(* Logix 5000 project; controller TFF vendor 1 type 14 code 107 rev 33.11; software revision 33.04; part 16 of 38 *)
(* tags used below, declared in another part *)
   AddressTotalizer : DINT;   // Temp Address used in modPhaseTotal
   Index : DINT;   // Index
   PLCDST : SINT;   // Current PLC Day Light Saving
   PLCTimeZoneString : STRING;   // Current PLC TimeZone
   TimeZoneUTC0 : STRING;   // String value for Time zone UTC 0
   AnalogPoint : AnalogInput[50];   // Analog Input Array
   Concentration : Concentration;
   ControlLoop_PCV101 : ALIAS FOR ControlLoop[3];
   ControlLoop_PCV101_5ms : ALIAS FOR ControlLoop[4];
   ControlLoop_PCV101_RAMP_OUT : REAL;   // Ramp Output
   Diafiltration : Diafiltration;
   FI201 : ALIAS FOR AnalogPoint[2];
   FQ_Conc : ALIAS FOR Totalizer[0];   // Concentration Totalizer
   FQ_Diaf : ALIAS FOR Totalizer[1];   // DiafiltrationTotalizer
   MiscREAL : REAL[50];   // Misc Real Values
   PCDateTime : DINT[7];   // Date/Time Array from PC
   PCV101 : ALIAS FOR AnalogPoint[3];
   PCV101_Control : PCV_Control;   // PCV101 Control UDT
   PCV101_PID : PCV;   // PCV101 PID Management
   Phase : Phases[6];   // Phase Control Array
   PhaseTotalizer : PhaseTotalizer[18];   // Phase Totalizers Array
   Rack_Murr_Node1_TFF20 : IO_Station;   // Status of Node 1 TFF20
   Rack_Murr_Node1_TFF40 : IO_Station;   // Status of Node 1 TFF40
   Rack_Murr_Node1_TFF80 : IO_Station;   // Status of Node 1 TFF80
   RawAnalogInputArray : INT[50];   // Array of analog input raw
   SysControl : SysControl;   // General system status and command
   ThisSystem : SystemType;
   TimerControl : TimerControl;   // Timer Control
   Timers : Timers[22];   // Timer Array
   Totalizer : Totalizers[20];   // Totalizers Array
   Valve : Valve[100];   // Valve Array
(* MainProgram, continued *)

ROUTINE modPhaseTotal   (* ladder *)
// Phase Totalizer Module
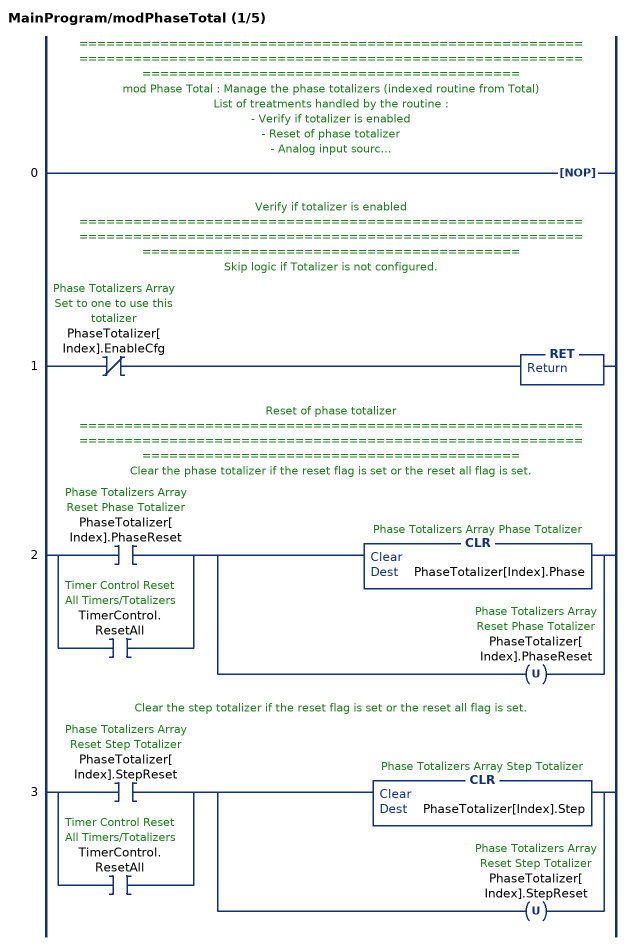
   // ==========================================================================================================================================================
   //                                                                                                   mod Phase Total : Manage the phase totalizers (indexed routine from Total)
   //                                                     List of treatments handled by the routine :
   //                                                          - Verify if totalizer is enabled
   //                                                          - Reset of phase totalizer
   //                                                          - Analog input source
   //                                                          - Calculating the totalizer values
   //                                                     -----------------------------------------------------------------------------------------------------------------------------------------------------
   //                                                     History
   // 		2019-DEC-24 - Merck - Q. Spindler - Initial version for Candidate Release 1.00.00.00.a
   // ==========================================================================================================================================================
   0: NOP();
   // Verify if totalizer is enabled
   // ==========================================================================================================================================================
   // Skip logic if Totalizer is not configured.
   1: XIO(PhaseTotalizer[Index].EnableCfg)RET();
   // Reset of phase totalizer
   // ==========================================================================================================================================================
   // Clear the phase totalizer if the reset flag is set or the reset all flag is set.
   2: [XIC(PhaseTotalizer[Index].PhaseReset) ,XIC(TimerControl.ResetAll) ][CLR(PhaseTotalizer[Index].Phase) ,OTU(PhaseTotalizer[Index].PhaseReset) ];
   // Clear the step totalizer if the reset flag is set or the reset all flag is set.
   3: [XIC(PhaseTotalizer[Index].StepReset) ,XIC(TimerControl.ResetAll) ][CLR(PhaseTotalizer[Index].Step) ,OTU(PhaseTotalizer[Index].StepReset) ];
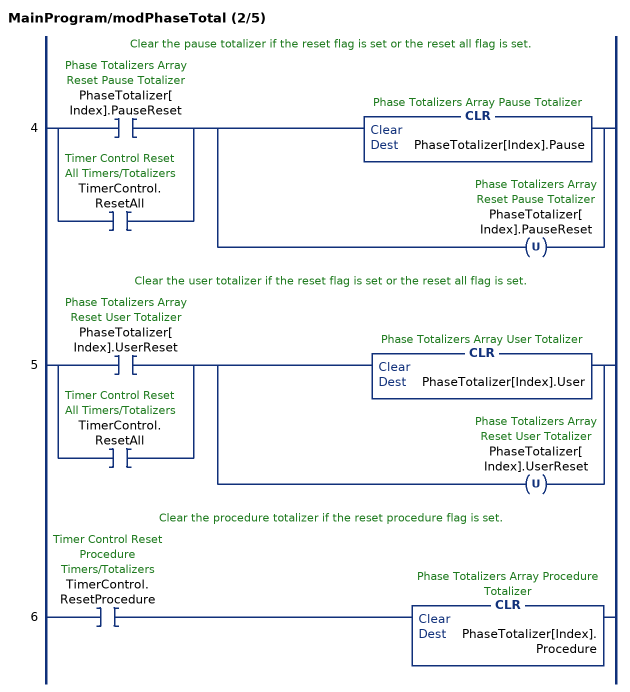
   // Clear the pause totalizer if the reset flag is set or the reset all flag is set.
   4: [XIC(PhaseTotalizer[Index].PauseReset) ,XIC(TimerControl.ResetAll) ][CLR(PhaseTotalizer[Index].Pause) ,OTU(PhaseTotalizer[Index].PauseReset) ];
   // Clear the user totalizer if the reset flag is set or the reset all flag is set.
   5: [XIC(PhaseTotalizer[Index].UserReset) ,XIC(TimerControl.ResetAll) ][CLR(PhaseTotalizer[Index].User) ,OTU(PhaseTotalizer[Index].UserReset) ];
   // Clear the procedure totalizer if the reset procedure flag is set.
   6: XIC(TimerControl.ResetProcedure)CLR(PhaseTotalizer[Index].Procedure);
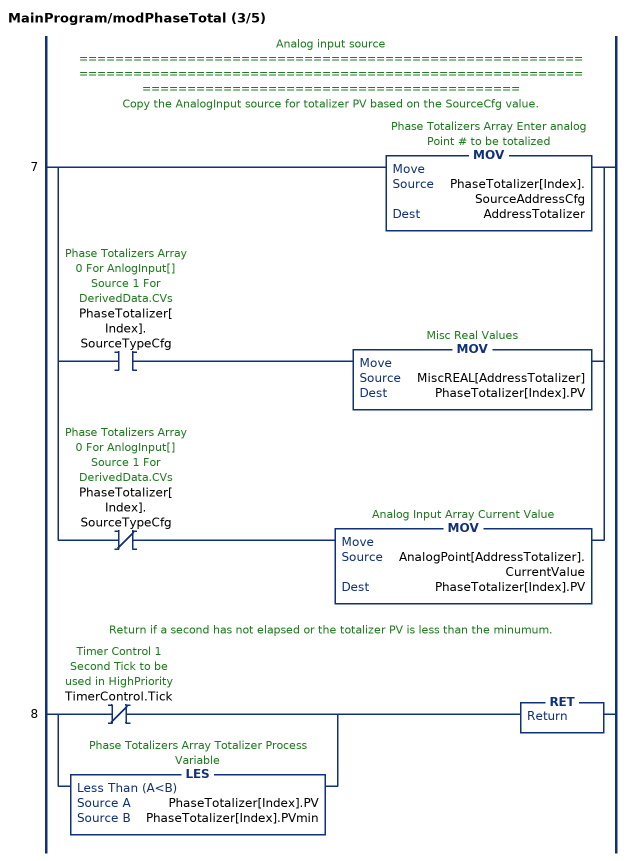
   // Analog input source
   // ==========================================================================================================================================================
   // Copy the AnalogInput source for totalizer PV based on the SourceCfg value.
   7: [MOV(PhaseTotalizer[Index].SourceAddressCfg,AddressTotalizer) ,XIC(PhaseTotalizer[Index].SourceTypeCfg) MOV(MiscREAL[AddressTotalizer],PhaseTotalizer[Index].PV) ,XIO(PhaseTotalizer[Index].SourceTypeCfg) MOV(AnalogPoint[AddressTotalizer].CurrentValue,PhaseTotalizer[Index].PV) ];
   // Return if a second has not elapsed or the totalizer PV is less than the minumum.
   8: [XIO(TimerControl.Tick) ,LES(PhaseTotalizer[Index].PV,PhaseTotalizer[Index].PVmin) ]RET();
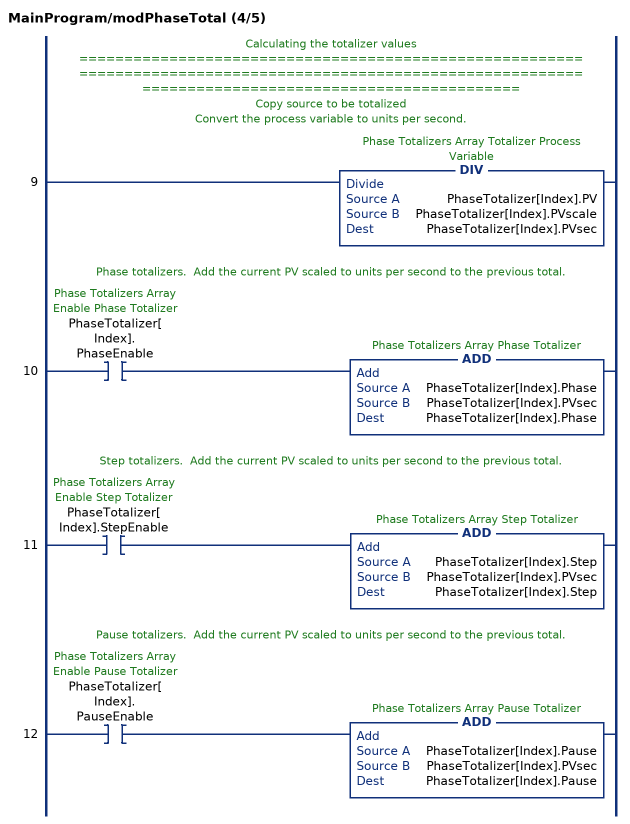
   // Calculating the totalizer values
   // ==========================================================================================================================================================
   // Copy source to be totalized
   // Convert the process variable to units per second.
   9: DIV(PhaseTotalizer[Index].PV,PhaseTotalizer[Index].PVscale,PhaseTotalizer[Index].PVsec);
   // Phase totalizers.  Add the current PV scaled to units per second to the previous total.
   10: XIC(PhaseTotalizer[Index].PhaseEnable)ADD(PhaseTotalizer[Index].Phase,PhaseTotalizer[Index].PVsec,PhaseTotalizer[Index].Phase);
   // Step totalizers.  Add the current PV scaled to units per second to the previous total.
   11: XIC(PhaseTotalizer[Index].StepEnable)ADD(PhaseTotalizer[Index].Step,PhaseTotalizer[Index].PVsec,PhaseTotalizer[Index].Step);
   // Pause totalizers.  Add the current PV scaled to units per second to the previous total.
   12: XIC(PhaseTotalizer[Index].PauseEnable)ADD(PhaseTotalizer[Index].Pause,PhaseTotalizer[Index].PVsec,PhaseTotalizer[Index].Pause);
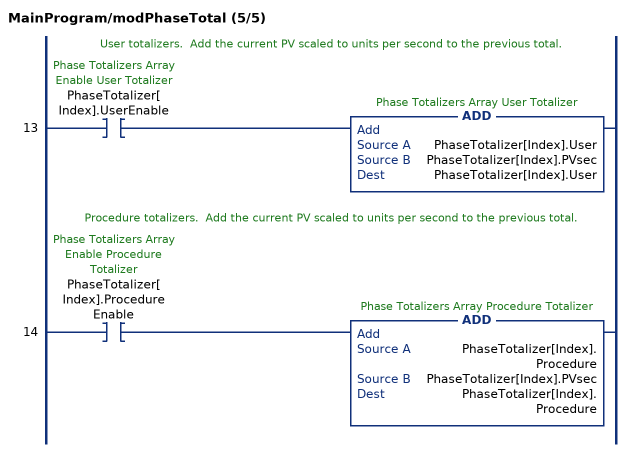
   // User totalizers.  Add the current PV scaled to units per second to the previous total.
   13: XIC(PhaseTotalizer[Index].UserEnable)ADD(PhaseTotalizer[Index].User,PhaseTotalizer[Index].PVsec,PhaseTotalizer[Index].User);
   // Procedure totalizers.  Add the current PV scaled to units per second to the previous total.
   14: XIC(PhaseTotalizer[Index].ProcedureEnable)ADD(PhaseTotalizer[Index].Procedure,PhaseTotalizer[Index].PVsec,PhaseTotalizer[Index].Procedure);
END_ROUTINE

ROUTINE modTotal   (* ladder *)
// Totalizer Module
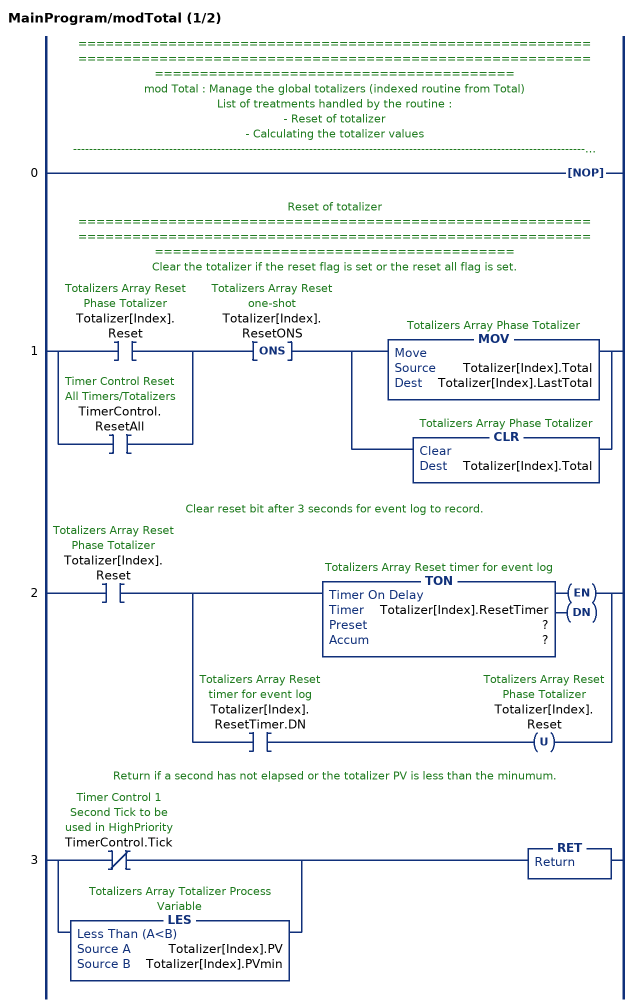
   // ==========================================================================================================================================================
   //                                                                                                   mod Total : Manage the global totalizers (indexed routine from Total)
   //                                                     List of treatments handled by the routine :
   //                                                          - Reset of totalizer
   //                                                          - Calculating the totalizer values
   //                                                     -----------------------------------------------------------------------------------------------------------------------------------------------------
   //                                                     History
   // 		2019-DEC-24 - Merck - Q. Spindler - Initial version for Candidate Release 1.00.00.00.a
   // ==========================================================================================================================================================
   0: NOP();
   // Reset of totalizer
   // ==========================================================================================================================================================
   // Clear the totalizer if the reset flag is set or the reset all flag is set.
   1: [XIC(Totalizer[Index].Reset) ,XIC(TimerControl.ResetAll) ]ONS(Totalizer[Index].ResetONS)[MOV(Totalizer[Index].Total,Totalizer[Index].LastTotal) ,CLR(Totalizer[Index].Total) ];
   // Clear reset bit after 3 seconds for event log to record.
   2: XIC(Totalizer[Index].Reset)[TON(Totalizer[Index].ResetTimer,?,?) ,XIC(Totalizer[Index].ResetTimer.DN) OTU(Totalizer[Index].Reset) ];
   // Return if a second has not elapsed or the totalizer PV is less than the minumum.
   3: [XIO(TimerControl.Tick) ,LES(Totalizer[Index].PV,Totalizer[Index].PVmin) ]RET();
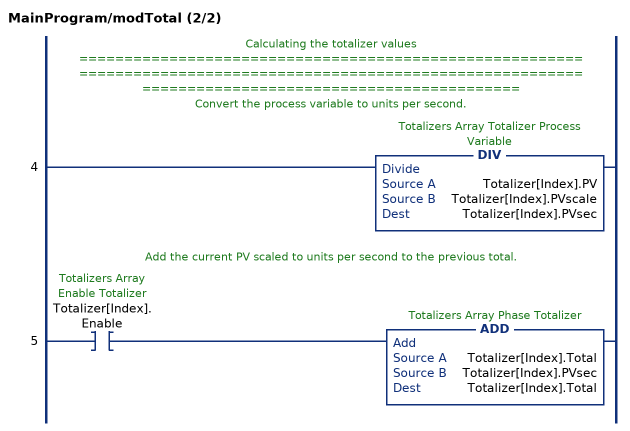
   // Calculating the totalizer values
   // ==========================================================================================================================================================
   // Convert the process variable to units per second.
   4: DIV(Totalizer[Index].PV,Totalizer[Index].PVscale,Totalizer[Index].PVsec);
   // Add the current PV scaled to units per second to the previous total.
   5: XIC(Totalizer[Index].Enable)ADD(Totalizer[Index].Total,Totalizer[Index].PVsec,Totalizer[Index].Total);
END_ROUTINE

ROUTINE PCDateTime   (* structured text *)
   (* =======================================================================
   	PCDateTime : Synchronize the PLC with PC clock
   
   	List of treatments
   		- Synchronization
   
   -----------------------------------------------------------------------------------------------------------------------------------------------------
   	History
   		2019-DEC-24 - Merck - Q. Spindler - Initial version for Candidate Release 1.00.00.00.a
   =========================================================================*)
   
   
   (* Synchronization
   =========================================================================*)
   (*Update the internal PLC clock with the PC clock when the microseconds value is not -1*)
   IF PCDateTime[6] <> -1 THEN;
   	SSV (WALLCLOCKTIME, , DateTime, PCDateTime[0]);
   	PCDateTime[6] := -1;
   END_IF;
   
   (*Get PLC DST settings and set it to 0 of not already*)
   GSV (WALLCLOCKTIME, ,ApplyDST , PLCDST);
   IF PLCDST <> 0 THEN;
   	PLCDST := 0;
   	SSV (WALLCLOCKTIME, ,ApplyDST , PLCDST);
   END_IF;
   
   (*Get PLC TimeZone and set it to UTC0 of not already*)
   GSV (WALLCLOCKTIME, ,TimeZoneString, PLCTimeZoneString);
   IF PLCTimeZoneString <> TimeZoneUTC0 THEN;
   	SSV (WALLCLOCKTIME, ,TimeZoneString , TimeZoneUTC0);
   END_IF;
   
END_ROUTINE

ROUTINE Time   (* ladder *)
// Timekeeping Routine
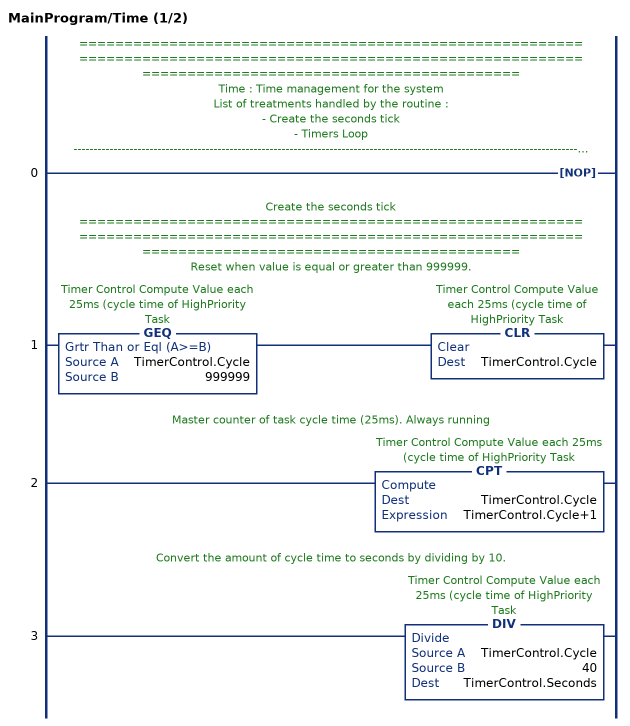
   // ==========================================================================================================================================================
   //                                                                                                                       Time : Time management for the system
   //                                                     List of treatments handled by the routine :
   //                                                          - Create the seconds tick
   //                                                          - Timers Loop
   //                                                     -----------------------------------------------------------------------------------------------------------------------------------------------------
   //                                                     History
   // 		2019-DEC-24 - Merck - Q. Spindler - Initial version for Candidate Release 1.00.00.00.a
   //                                 2020-APR-06 - Merck - Q. Spindler - Modifications for Candidate Release 1.00.00.00.b
   // Add TimerControl.NewTickMainTask
   // ==========================================================================================================================================================
   0: NOP();
   // Create the seconds tick
   // ==========================================================================================================================================================
   // Reset when value is equal or greater than 999999.
   1: GEQ(TimerControl.Cycle,999999)CLR(TimerControl.Cycle);
   // Master counter of task cycle time (25ms). Always running
   2: CPT(TimerControl.Cycle,TimerControl.Cycle+1);
   // Convert the amount of cycle time to seconds by dividing by 10.
   3: DIV(TimerControl.Cycle,40,TimerControl.Seconds);
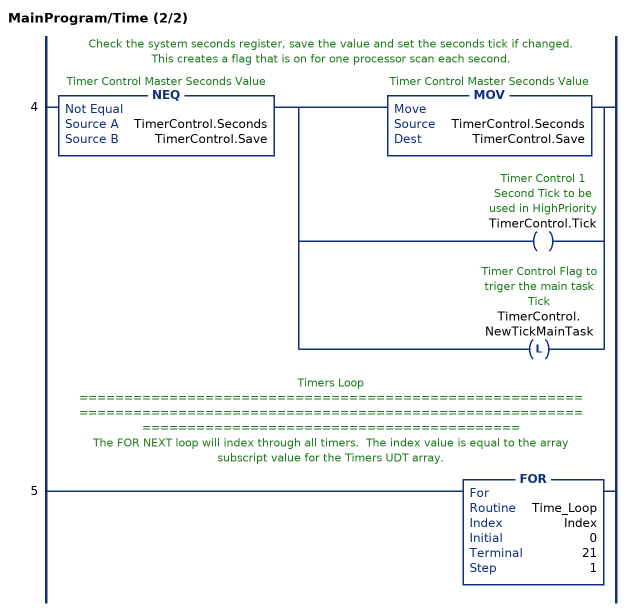
   // Check the system seconds register, save the value and set the seconds tick if changed.  This creates a flag that is on for one processor scan each second.
   4: NEQ(TimerControl.Seconds,TimerControl.Save)[MOV(TimerControl.Seconds,TimerControl.Save) ,OTE(TimerControl.Tick) ,OTL(TimerControl.NewTickMainTask) ];
   // Timers Loop
   // ==========================================================================================================================================================
   // The FOR NEXT loop will index through all timers.  The index value is equal to the array subscript value for the Timers UDT array.
   5: FOR(Time_Loop,Index,0,21,1);
END_ROUTINE

ROUTINE Time_Loop   (* ladder *)
// Timer Routine
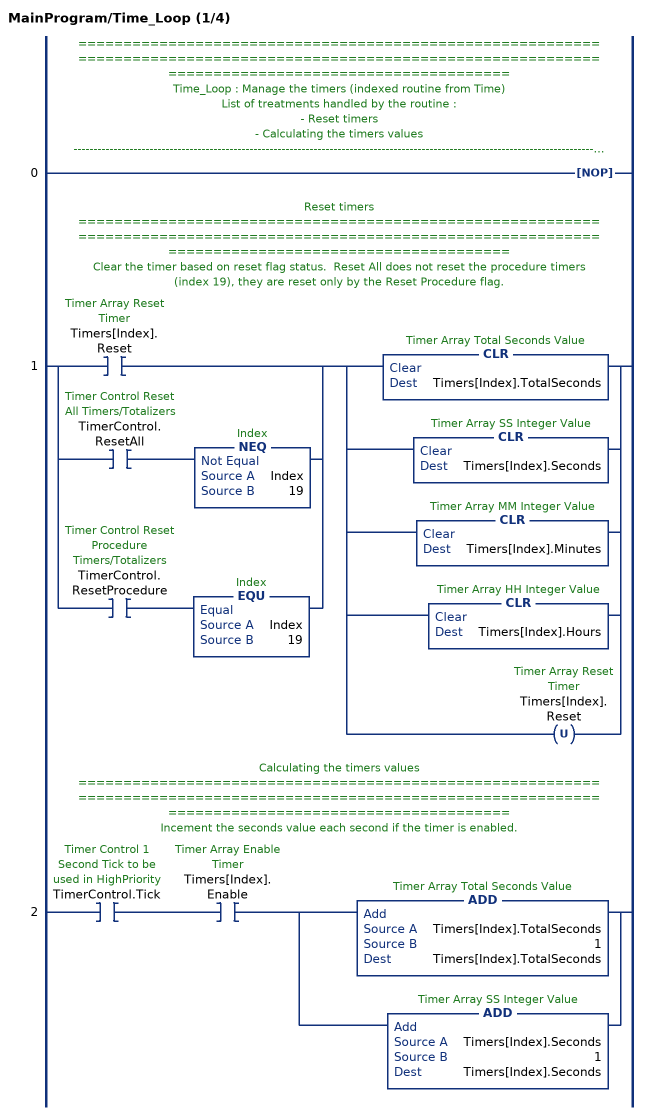
   // ==========================================================================================================================================================
   //                                                                                                              Time_Loop : Manage the timers (indexed routine from Time)
   //                                                     List of treatments handled by the routine :
   //                                                          - Reset timers
   //                                                          - Calculating the timers values
   //                                                     -----------------------------------------------------------------------------------------------------------------------------------------------------
   //                                                     History
   // 		2019-DEC-24 - Merck - Q. Spindler - Initial version for Candidate Release 1.00.00.00.a
   // ==========================================================================================================================================================
   0: NOP();
   // Reset timers
   // ==========================================================================================================================================================
   // Clear the timer based on reset flag status.  Reset All does not reset the procedure timers (index 19), they are reset only by the Reset Procedure flag.
   1: [XIC(Timers[Index].Reset) ,XIC(TimerControl.ResetAll) NEQ(Index,19) ,XIC(TimerControl.ResetProcedure) EQU(Index,19) ][CLR(Timers[Index].TotalSeconds) ,CLR(Timers[Index].Seconds) ,CLR(Timers[Index].Minutes) ,CLR(Timers[Index].Hours) ,OTU(Timers[Index].Reset) ];
   // Calculating the timers values
   // ==========================================================================================================================================================
   // Incement the seconds value each second if the timer is enabled.
   2: XIC(TimerControl.Tick)XIC(Timers[Index].Enable)[ADD(Timers[Index].TotalSeconds,1,Timers[Index].TotalSeconds) ,ADD(Timers[Index].Seconds,1,Timers[Index].Seconds) ];
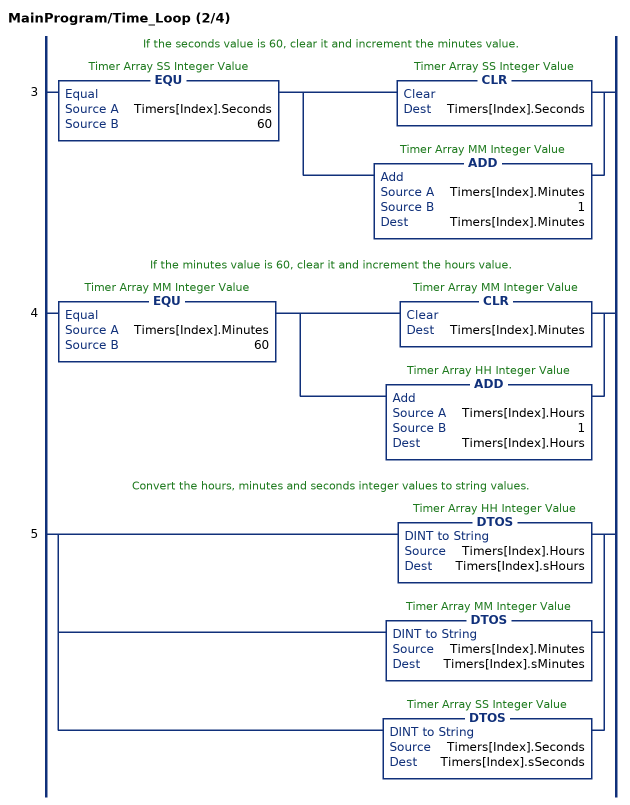
   // If the seconds value is 60, clear it and increment the minutes value.
   3: EQU(Timers[Index].Seconds,60)[CLR(Timers[Index].Seconds) ,ADD(Timers[Index].Minutes,1,Timers[Index].Minutes) ];
   // If the minutes value is 60, clear it and increment the hours value.
   4: EQU(Timers[Index].Minutes,60)[CLR(Timers[Index].Minutes) ,ADD(Timers[Index].Hours,1,Timers[Index].Hours) ];
   // Convert the hours, minutes and seconds integer values to string values.
   5: [DTOS(Timers[Index].Hours,Timers[Index].sHours) ,DTOS(Timers[Index].Minutes,Timers[Index].sMinutes) ,DTOS(Timers[Index].Seconds,Timers[Index].sSeconds) ];
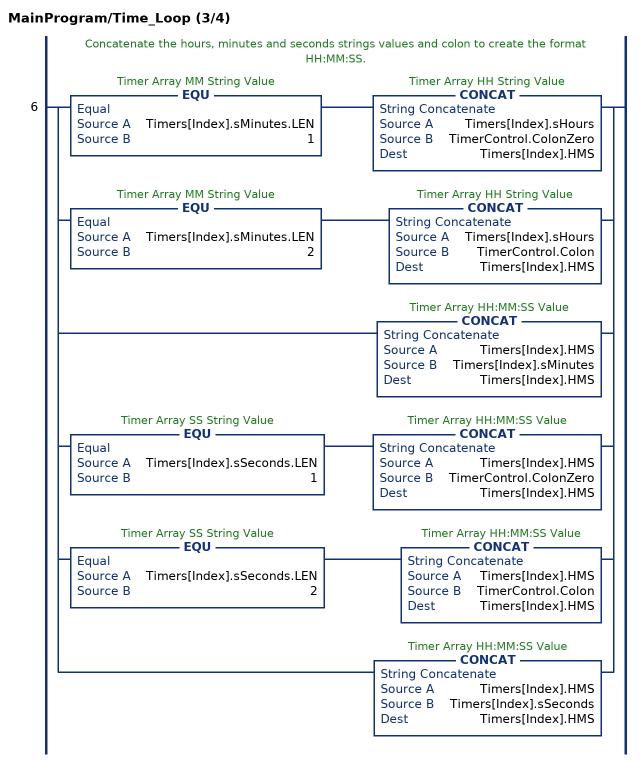
   // Concatenate the hours, minutes and seconds strings values and colon to create the format HH:MM:SS.
   6: [EQU(Timers[Index].sMinutes.LEN,1) CONCAT(Timers[Index].sHours,TimerControl.ColonZero,Timers[Index].HMS) ,EQU(Timers[Index].sMinutes.LEN,2) CONCAT(Timers[Index].sHours,TimerControl.Colon,Timers[Index].HMS) ,CONCAT(Timers[Index].HMS,Timers[Index].sMinutes,Timers[Index].HMS) ,EQU(Timers[Index].sSeconds.LEN,1) CONCAT(Timers[Index].HMS,TimerControl.ColonZero,Timers[Index].HMS) ,EQU(Timers[Index].sSeconds.LEN,2) CONCAT(Timers[Index].HMS,TimerControl.Colon,Timers[Index].HMS) ,CONCAT(Timers[Index].HMS,Timers[Index].sSeconds,Timers[Index].HMS) ];
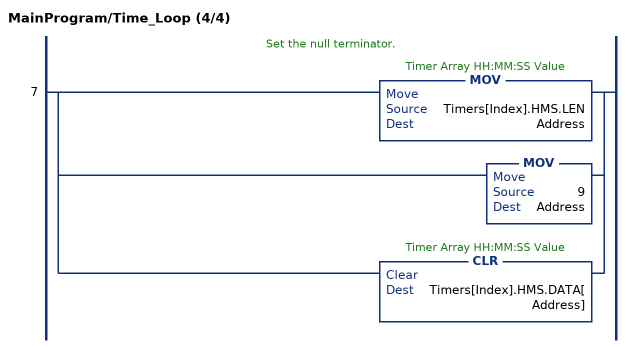
   // Set the null terminator.
   7: [[MOV(Timers[Index].HMS.LEN,Address) ,MOV(9,Address) ] ,CLR(Timers[Index].HMS.DATA[Address]) ];
END_ROUTINE

ROUTINE Total   (* ladder *)
// Totalizer Routine
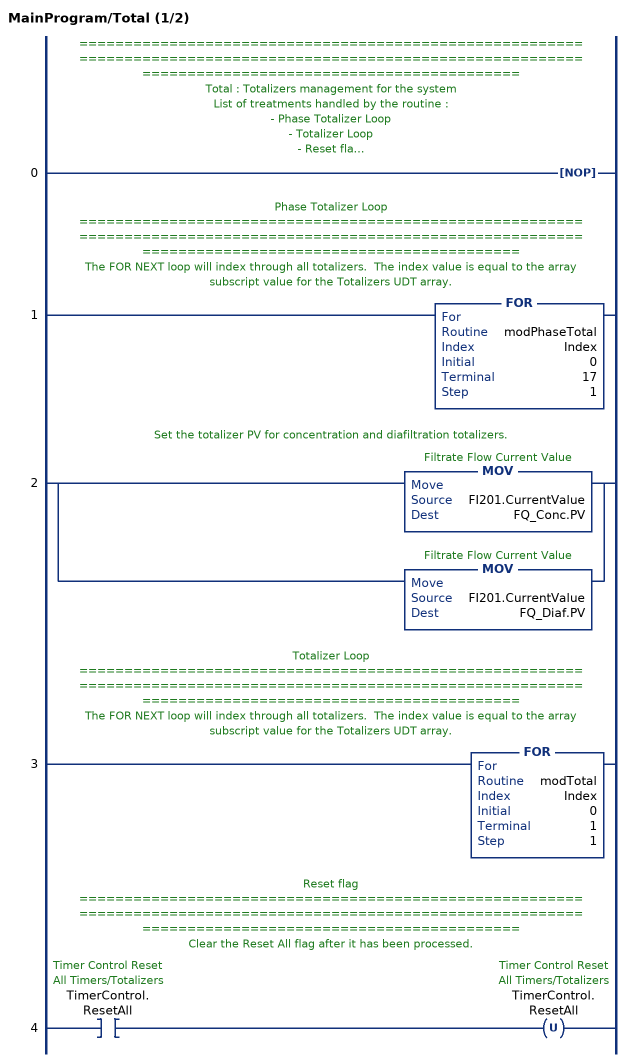
   // ==========================================================================================================================================================
   //                                                                                                              Total : Totalizers management for the system
   //                                                     List of treatments handled by the routine :
   //                                                          - Phase Totalizer Loop
   //                                                          - Totalizer Loop
   //                                                          - Reset flag
   //                                                     -----------------------------------------------------------------------------------------------------------------------------------------------------
   //                                                     History
   // 		2019-DEC-24 - Merck - Q. Spindler - Initial version for Candidate Release 1.00.00.00.a
   //                                2022-JAN-11 - Merck - Q. Spindler - Modifications for Candidate Release 1.01.00.00.a
   //   - Change Phase Totalizer size
   // ==========================================================================================================================================================
   0: NOP();
   // Phase Totalizer Loop
   // ==========================================================================================================================================================
   // The FOR NEXT loop will index through all totalizers.  The index value is equal to the array subscript value for the Totalizers UDT array.
   1: FOR(modPhaseTotal,Index,0,17,1);
   // Set the totalizer PV for concentration and diafiltration totalizers.
   2: [MOV(FI201.CurrentValue,FQ_Conc.PV) ,MOV(FI201.CurrentValue,FQ_Diaf.PV) ];
   // Totalizer Loop
   // ==========================================================================================================================================================
   // The FOR NEXT loop will index through all totalizers.  The index value is equal to the array subscript value for the Totalizers UDT array.
   3: FOR(modTotal,Index,0,1,1);
   // Reset flag
   // ==========================================================================================================================================================
   // Clear the Reset All flag after it has been processed.
   4: XIC(TimerControl.ResetAll)OTU(TimerControl.ResetAll);
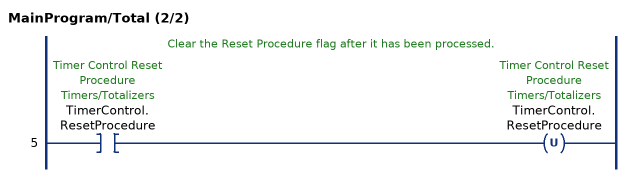
   // Clear the Reset Procedure flag after it has been processed.
   5: XIC(TimerControl.ResetProcedure)OTU(TimerControl.ResetProcedure);
END_ROUTINE
END_PROGRAM

PROGRAM MainProgram5ms   (* main routine MainRoutine, fault routine FaultRoutine *)
VAR
   Address : DINT := 1;   // Index
   Address2 : DINT := 41;
   ONS_PID02 : BOOL;
   PCV001_PID_Settings : INT;
   PCV101_AutoMaxRate : REAL := 0.25;   // PCV101 Maximum Rate in Auto Mode
   PCV101_ManualMaxRate : REAL := 0.01;   // PCV101 Maximum Rate in Manual mode
   PCV101_Max_CV : REAL := 100.01;   // Max CV for PCV101
   PCV101_PID_Settings : INT;
   SCL : SCALE := (InRawMax := 32767.0, InRawMin := 6553.0, InEUMax := 2000.0, Out := -499.96185, MinAlarm := 1);   // Scale Function
END_VAR

ROUTINE Control_Loop_PCV101_5ms   (* ladder *)
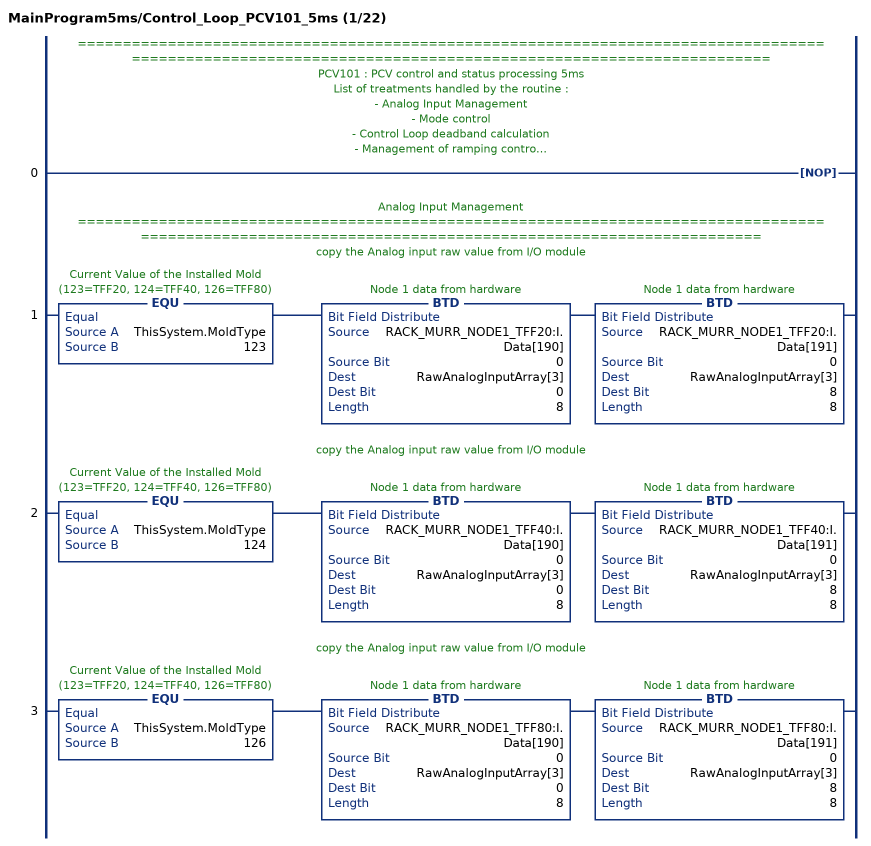
   // ==========================================================================================================================================================
   //                                                  PCV101 : PCV control and status processing 5ms
   //                                                     List of treatments handled by the routine :
   //                                                          - Analog Input Management
   //                                                          - Mode control
   //                                                          - Control Loop deadband calculation
   //                                                          - Management of ramping control
   //                                                          - Management of PID instruction
   //                                                          - PCV101 Control Valve Calibration
   //                                                          - Control of the analog output
   //                                                          - Loop status for HMI
   //                                                     -----------------------------------------------------------------------------------------------------------------------------------------------------
   //                                                     History
   // 		2019-DEC-24 - Merck - Q. Spindler - Initial version for Candidate Release 1.00.00.00.a
   // 		2021-APR-19 - Merck - Q. Spindler - Modifications for Candidate Release 1.00.00.00.e
   //                              - Add limit for the Output if greater than the Maximum CV
   //                                     - Add Compute the Maximum CV based on the Maximum Rate
   //                                                    - Start the PCV to close at 550 point instead of 0 (a bit less than 2 bar)
   // ==========================================================================================================================================================
   0: NOP();
   // Analog Input Management
   // ========================================================================================================================================================
   // copy the Analog input raw value from I/O module
   1: EQU(ThisSystem.MoldType,123)BTD(RACK_MURR_NODE1_TFF20:I.Data[190],0,RawAnalogInputArray[3],0,8)BTD(RACK_MURR_NODE1_TFF20:I.Data[191],0,RawAnalogInputArray[3],8,8);
   // copy the Analog input raw value from I/O module
   2: EQU(ThisSystem.MoldType,124)BTD(RACK_MURR_NODE1_TFF40:I.Data[190],0,RawAnalogInputArray[3],0,8)BTD(RACK_MURR_NODE1_TFF40:I.Data[191],0,RawAnalogInputArray[3],8,8);
   // copy the Analog input raw value from I/O module
   3: EQU(ThisSystem.MoldType,126)BTD(RACK_MURR_NODE1_TFF80:I.Data[190],0,RawAnalogInputArray[3],0,8)BTD(RACK_MURR_NODE1_TFF80:I.Data[191],0,RawAnalogInputArray[3],8,8);
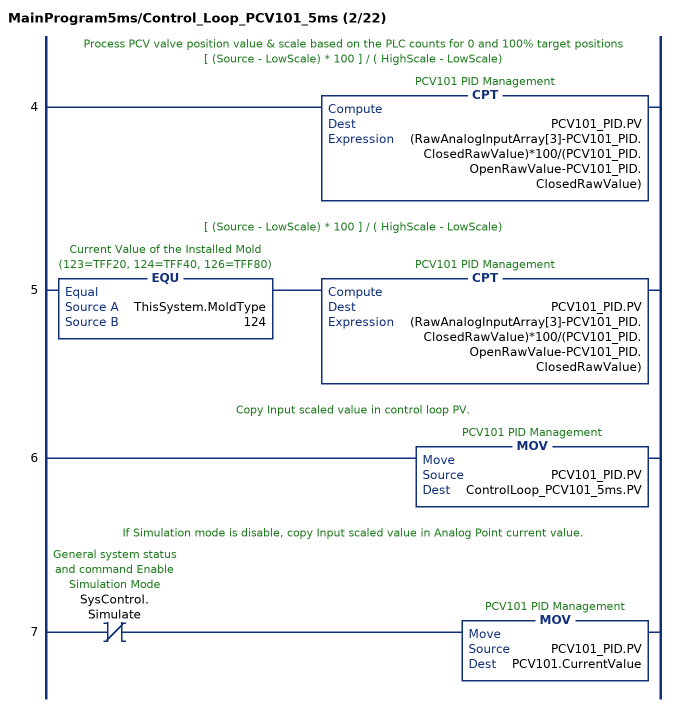
   // Process PCV valve position value & scale based on the PLC counts for 0 and 100% target positions
   // [ (Source - LowScale) * 100 ] / ( HighScale - LowScale)
   4: CPT(PCV101_PID.PV,(RawAnalogInputArray[3]-PCV101_PID.ClosedRawValue)*100/(PCV101_PID.OpenRawValue-PCV101_PID.ClosedRawValue));
   // [ (Source - LowScale) * 100 ] / ( HighScale - LowScale)
   5: EQU(ThisSystem.MoldType,124)CPT(PCV101_PID.PV,(RawAnalogInputArray[3]-PCV101_PID.ClosedRawValue)*100/(PCV101_PID.OpenRawValue-PCV101_PID.ClosedRawValue));
   // Copy Input scaled value in control loop PV.
   6: MOV(PCV101_PID.PV,ControlLoop_PCV101_5ms.PV);
   // If Simulation mode is disable, copy Input scaled value in Analog Point current value.
   7: XIO(SysControl.Simulate)MOV(PCV101_PID.PV,PCV101.CurrentValue);
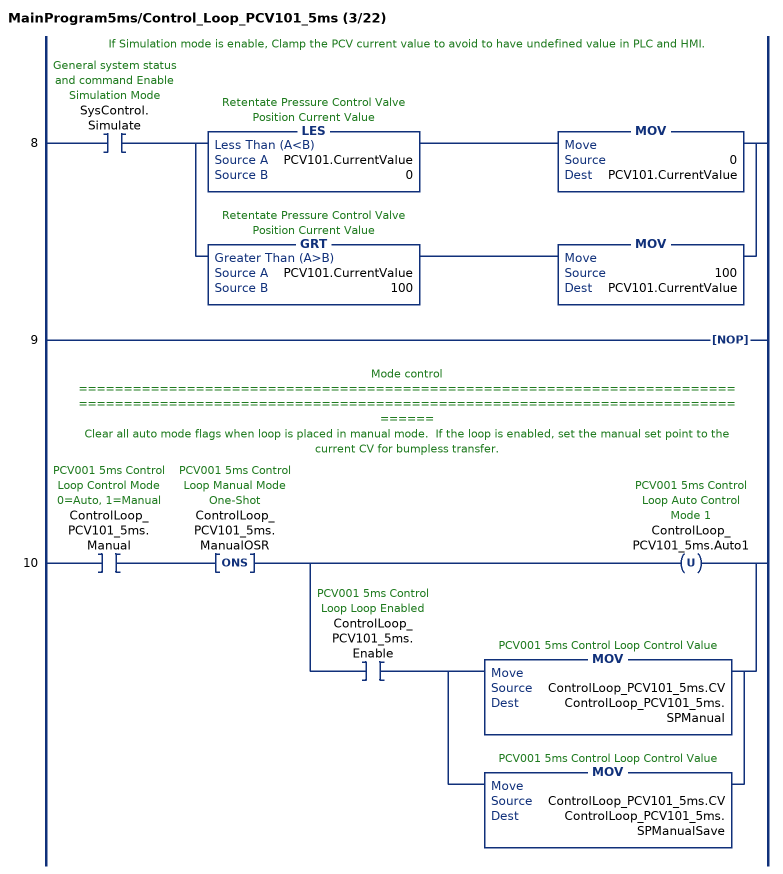
   // If Simulation mode is enable, Clamp the PCV current value to avoid to have undefined value in PLC and HMI.
   8: XIC(SysControl.Simulate)[LES(PCV101.CurrentValue,0) MOV(0,PCV101.CurrentValue) ,GRT(PCV101.CurrentValue,100) MOV(100,PCV101.CurrentValue) ];
   9: NOP();
   // Mode control
   // ========================================================================================================================================================
   // Clear all auto mode flags when loop is placed in manual mode.  If the loop is enabled, set the manual set point to the current CV for bumpless transfer.
   10: XIC(ControlLoop_PCV101_5ms.Manual)ONS(ControlLoop_PCV101_5ms.ManualOSR)[OTU(ControlLoop_PCV101_5ms.Auto1) ,XIC(ControlLoop_PCV101_5ms.Enable) [MOV(ControlLoop_PCV101_5ms.CV,ControlLoop_PCV101_5ms.SPManual) ,MOV(ControlLoop_PCV101_5ms.CV,ControlLoop_PCV101_5ms.SPManualSave) ] ];
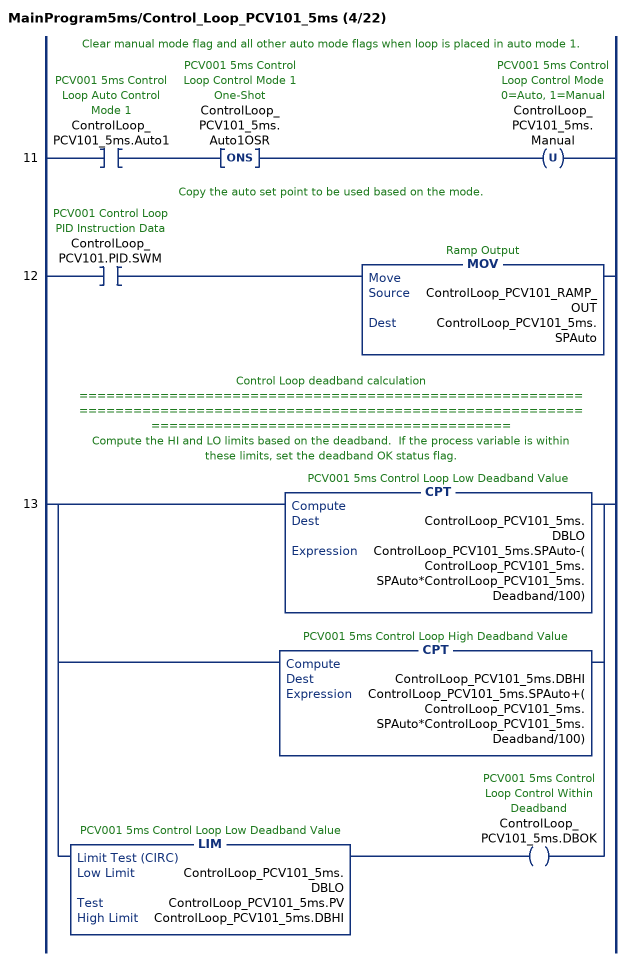
   // Clear manual mode flag and all other auto mode flags when loop is placed in auto mode 1.
   11: XIC(ControlLoop_PCV101_5ms.Auto1)ONS(ControlLoop_PCV101_5ms.Auto1OSR)OTU(ControlLoop_PCV101_5ms.Manual);
   // Copy the auto set point to be used based on the mode.
   12: XIC(ControlLoop_PCV101.PID.SWM)MOV(ControlLoop_PCV101_RAMP_OUT,ControlLoop_PCV101_5ms.SPAuto);
   // Control Loop deadband calculation
   // ========================================================================================================================================================
   // Compute the HI and LO limits based on the deadband.  If the process variable is within these limits, set the deadband OK status flag.
   13: [CPT(ControlLoop_PCV101_5ms.DBLO,ControlLoop_PCV101_5ms.SPAuto-(ControlLoop_PCV101_5ms.SPAuto*ControlLoop_PCV101_5ms.Deadband/100)) ,CPT(ControlLoop_PCV101_5ms.DBHI,ControlLoop_PCV101_5ms.SPAuto+(ControlLoop_PCV101_5ms.SPAuto*ControlLoop_PCV101_5ms.Deadband/100)) ,LIM(ControlLoop_PCV101_5ms.DBLO,ControlLoop_PCV101_5ms.PV,ControlLoop_PCV101_5ms.DBHI) OTE(ControlLoop_PCV101_5ms.DBOK) ];
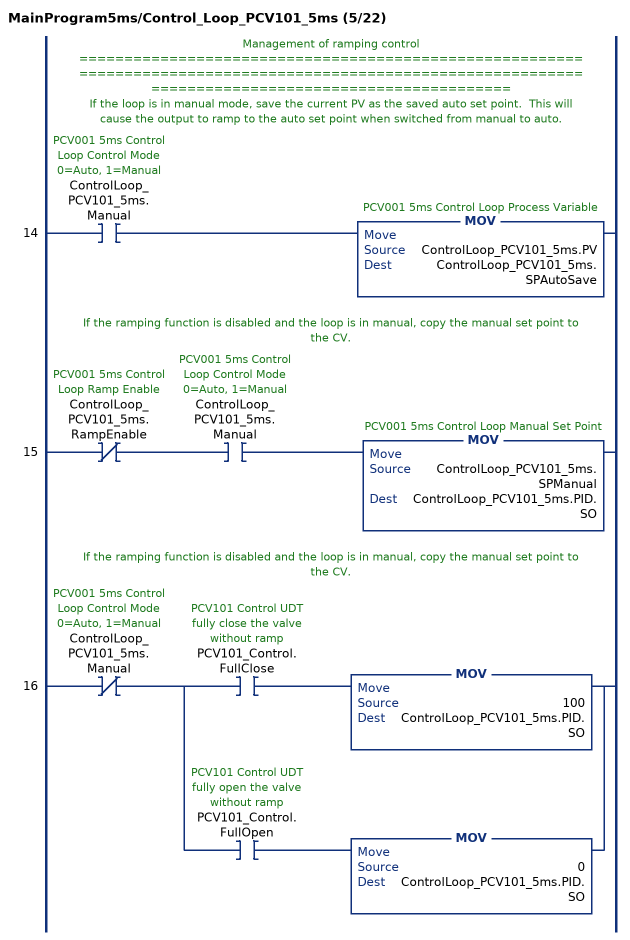
   // Management of ramping control
   // ========================================================================================================================================================
   // If the loop is in manual mode, save the current PV as the saved auto set point.  This will cause the output to ramp to the auto set point when switched from manual to auto.
   14: XIC(ControlLoop_PCV101_5ms.Manual)MOV(ControlLoop_PCV101_5ms.PV,ControlLoop_PCV101_5ms.SPAutoSave);
   // If the ramping function is disabled and the loop is in manual, copy the manual set point to the CV.
   15: XIO(ControlLoop_PCV101_5ms.RampEnable)XIC(ControlLoop_PCV101_5ms.Manual)MOV(ControlLoop_PCV101_5ms.SPManual,ControlLoop_PCV101_5ms.PID.SO);
   // If the ramping function is disabled and the loop is in manual, copy the manual set point to the CV.
   16: XIO(ControlLoop_PCV101_5ms.Manual)[XIC(PCV101_Control.FullClose) MOV(100,ControlLoop_PCV101_5ms.PID.SO) ,XIC(PCV101_Control.FullOpen) MOV(0,ControlLoop_PCV101_5ms.PID.SO) ];
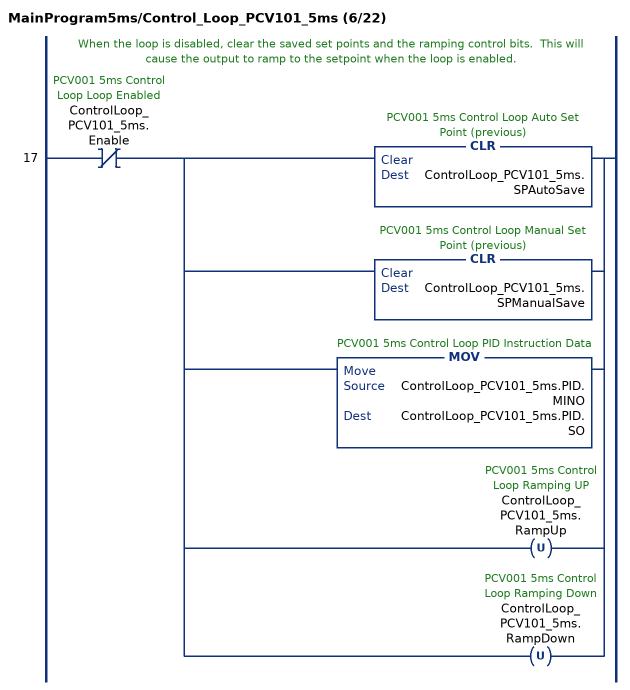
   // When the loop is disabled, clear the saved set points and the ramping control bits.  This will cause the output to ramp to the setpoint when the loop is enabled.
   17: XIO(ControlLoop_PCV101_5ms.Enable)[CLR(ControlLoop_PCV101_5ms.SPAutoSave) ,CLR(ControlLoop_PCV101_5ms.SPManualSave) ,MOV(ControlLoop_PCV101_5ms.PID.MINO,ControlLoop_PCV101_5ms.PID.SO) ,OTU(ControlLoop_PCV101_5ms.RampUp) ,OTU(ControlLoop_PCV101_5ms.RampDown) ];
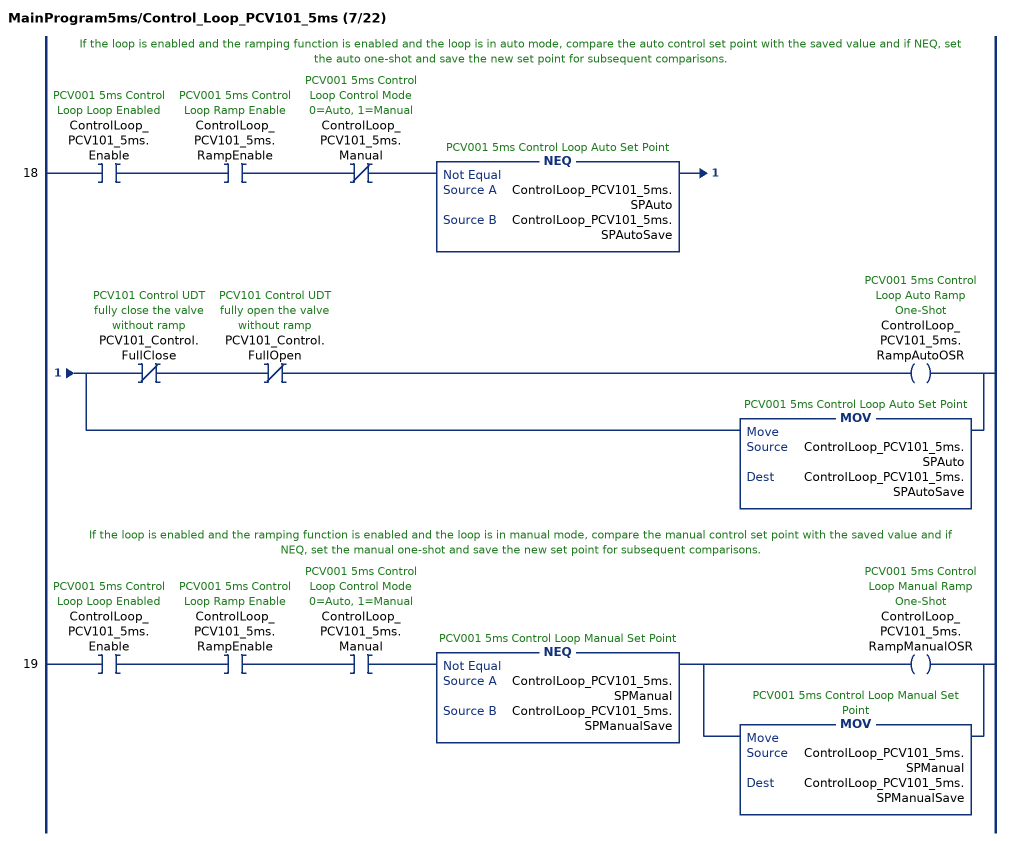
   // If the loop is enabled and the ramping function is enabled and the loop is in auto mode, compare the auto control set point with the saved value and if NEQ, set the auto one-shot and save the new set point for subsequent comparisons.
   18: XIC(ControlLoop_PCV101_5ms.Enable)XIC(ControlLoop_PCV101_5ms.RampEnable)XIO(ControlLoop_PCV101_5ms.Manual)NEQ(ControlLoop_PCV101_5ms.SPAuto,ControlLoop_PCV101_5ms.SPAutoSave)[XIO(PCV101_Control.FullClose) XIO(PCV101_Control.FullOpen) OTE(ControlLoop_PCV101_5ms.RampAutoOSR) ,MOV(ControlLoop_PCV101_5ms.SPAuto,ControlLoop_PCV101_5ms.SPAutoSave) ];
   // If the loop is enabled and the ramping function is enabled and the loop is in manual mode, compare the manual control set point with the saved value and if NEQ, set the manual one-shot and save the new set point for subsequent comparisons.
   19: XIC(ControlLoop_PCV101_5ms.Enable)XIC(ControlLoop_PCV101_5ms.RampEnable)XIC(ControlLoop_PCV101_5ms.Manual)NEQ(ControlLoop_PCV101_5ms.SPManual,ControlLoop_PCV101_5ms.SPManualSave)[OTE(ControlLoop_PCV101_5ms.RampManualOSR) ,MOV(ControlLoop_PCV101_5ms.SPManual,ControlLoop_PCV101_5ms.SPManualSave) ];
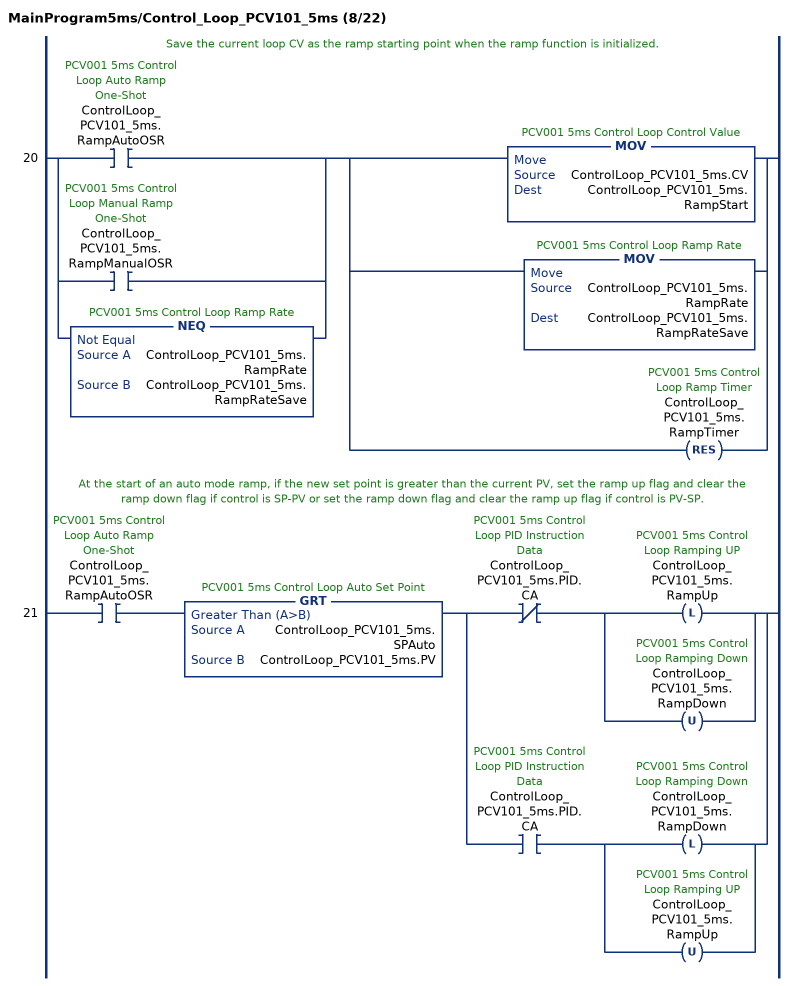
   // Save the current loop CV as the ramp starting point when the ramp function is initialized.
   20: [XIC(ControlLoop_PCV101_5ms.RampAutoOSR) ,XIC(ControlLoop_PCV101_5ms.RampManualOSR) ,NEQ(ControlLoop_PCV101_5ms.RampRate,ControlLoop_PCV101_5ms.RampRateSave) ][MOV(ControlLoop_PCV101_5ms.CV,ControlLoop_PCV101_5ms.RampStart) ,MOV(ControlLoop_PCV101_5ms.RampRate,ControlLoop_PCV101_5ms.RampRateSave) ,RES(ControlLoop_PCV101_5ms.RampTimer) ];
   // At the start of an auto mode ramp, if the new set point is greater than the current PV, set the ramp up flag and clear the ramp down flag if control is SP-PV or set the ramp down flag and clear the ramp up flag if control is PV-SP.
   21: XIC(ControlLoop_PCV101_5ms.RampAutoOSR)GRT(ControlLoop_PCV101_5ms.SPAuto,ControlLoop_PCV101_5ms.PV)[XIO(ControlLoop_PCV101_5ms.PID.CA) [OTL(ControlLoop_PCV101_5ms.RampUp) ,OTU(ControlLoop_PCV101_5ms.RampDown) ] ,XIC(ControlLoop_PCV101_5ms.PID.CA) [OTL(ControlLoop_PCV101_5ms.RampDown) ,OTU(ControlLoop_PCV101_5ms.RampUp) ] ];
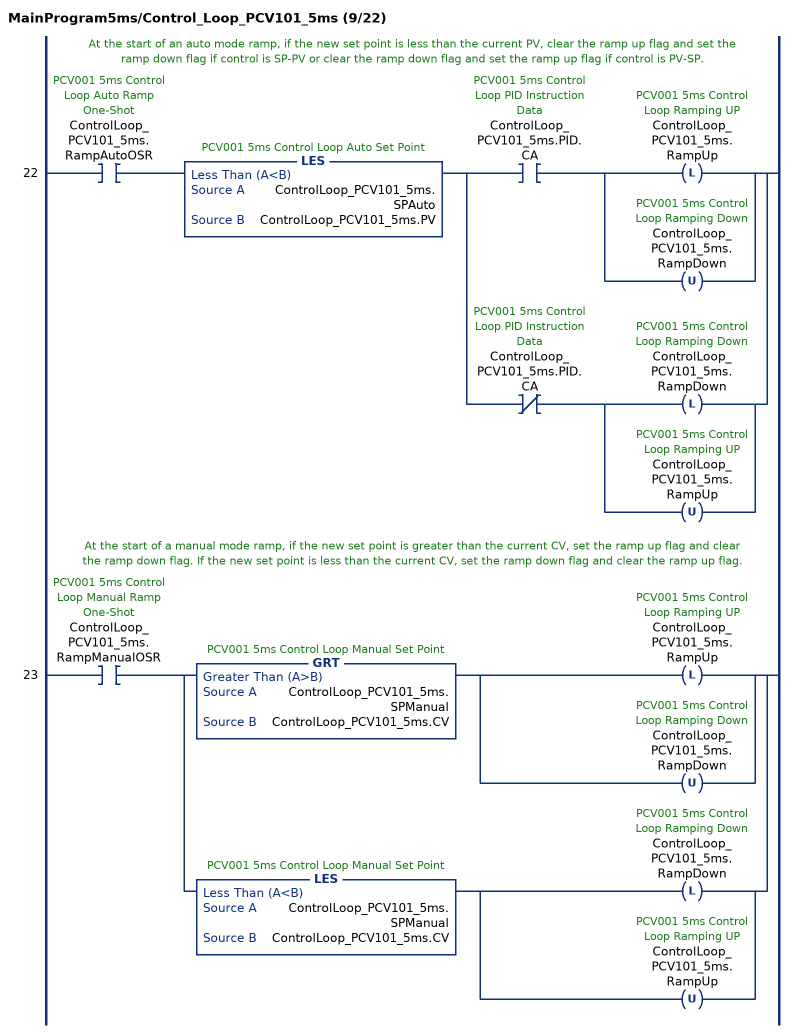
   // At the start of an auto mode ramp, if the new set point is less than the current PV, clear the ramp up flag and set the ramp down flag if control is SP-PV or clear the ramp down flag and set the ramp up flag if control is PV-SP.
   22: XIC(ControlLoop_PCV101_5ms.RampAutoOSR)LES(ControlLoop_PCV101_5ms.SPAuto,ControlLoop_PCV101_5ms.PV)[XIC(ControlLoop_PCV101_5ms.PID.CA) [OTL(ControlLoop_PCV101_5ms.RampUp) ,OTU(ControlLoop_PCV101_5ms.RampDown) ] ,XIO(ControlLoop_PCV101_5ms.PID.CA) [OTL(ControlLoop_PCV101_5ms.RampDown) ,OTU(ControlLoop_PCV101_5ms.RampUp) ] ];
   // At the start of a manual mode ramp, if the new set point is greater than the current CV, set the ramp up flag and clear the ramp down flag. If the new set point is less than the current CV, set the ramp down flag and clear the ramp up flag.
   23: XIC(ControlLoop_PCV101_5ms.RampManualOSR)[GRT(ControlLoop_PCV101_5ms.SPManual,ControlLoop_PCV101_5ms.CV) [OTL(ControlLoop_PCV101_5ms.RampUp) ,OTU(ControlLoop_PCV101_5ms.RampDown) ] ,LES(ControlLoop_PCV101_5ms.SPManual,ControlLoop_PCV101_5ms.CV) [OTL(ControlLoop_PCV101_5ms.RampDown) ,OTU(ControlLoop_PCV101_5ms.RampUp) ] ];
